// TIA Portal V18 export
TYPE "Modezone_Gap"
   STRUCT
      GapActive : Bool;
   END_STRUCT;
END_TYPE
